{attribute 'qualified_only'}
{attribute 'strict'}
TYPE ENUM_CurrentState :
(
	CloseValve := 0,
	OpenValve:=1,
	CirculateWater:=2,
	InsertPowder:=3
);
END_TYPE

(* stored: Version 1.1.0.1, ProductVersion 3.1.4024.12
   DUT ENUM_CurrentState: Id {ce786795-a470-4e9c-925e-e3435531e3ef} *)
